FUNCTION_BLOCK T_SafeSr_Tests EXTENDS TcUnit.FB_TestSuite
VAR
    // Test_SetDominantLatch
    group_1 : T_SafeGroup;
    fb_1 : T_SafeSr(group := group_1);
    // Test_UnconnectedResetIsRefused
    group_2 : T_SafeGroup;
    fb_2 : T_SafeSr(group := group_2);
END_VAR

Test_SetDominantLatch();
Test_UnconnectedResetIsRefused();

METHOD PRIVATE Test_SetDominantLatch
TcUnit.TEST(__POUNAME());
// act / assert
group_1(Run := TRUE);
fb_1(Set := TRUE, Reset := TRUE);
AssertEquals_BOOL(Expected := TRUE, Actual := fb_1.SrOut, Message := 'set dominant');
fb_1(Set := FALSE, Reset := TRUE);
AssertEquals_BOOL(Expected := FALSE, Actual := fb_1.SrOut, Message := 'reset');
fb_1(Set := FALSE, Reset := FALSE);
AssertEquals_BOOL(Expected := FALSE, Actual := fb_1.SrOut, Message := 'held');
TEST_FINISHED_NAMED(__POUNAME());
END_METHOD

METHOD PRIVATE Test_UnconnectedResetIsRefused
TcUnit.TEST(__POUNAME());
// arrange / act: Reset is unconnected, which the Safety Editor refuses
group_2(Run := TRUE);
fb_2(Set := TRUE);
group_2(Run := TRUE);
fb_2(Set := TRUE);
// assert
AssertEquals_BOOL(Expected := TRUE, Actual := fb_2.Error, Message := 'configuration error reported');
AssertEquals_BYTE(Expected := TO_BYTE(E_SafeFbState.Error), Actual := fb_2.State, Message := 'state ERROR');
AssertEquals_WORD(Expected := WORD#16#8000, Actual := fb_2.Diag, Message := 'diag bit 15 configuration refused');
AssertEquals_BOOL(Expected := FALSE, Actual := fb_2.SrOut, Message := 'SrOut stays at its safe value');
AssertEquals_BOOL(Expected := TRUE, Actual := group_2.FbErr, Message := 'the group sees an FB error');
// act: ErrAck 0 -> 1 -> 0 does not clear a configuration error
group_2(Run := TRUE, ErrAck := TRUE);
fb_2(Set := TRUE);
group_2(Run := TRUE, ErrAck := TRUE);
fb_2(Set := TRUE);
group_2(Run := TRUE, ErrAck := FALSE);
fb_2(Set := TRUE);
AssertEquals_BOOL(Expected := TRUE, Actual := fb_2.Error, Message := 'error not acknowledged');
AssertEquals_WORD(Expected := WORD#16#8000, Actual := fb_2.Diag, Message := 'diag bit 15 kept');
TEST_FINISHED_NAMED(__POUNAME());
END_METHOD

END_FUNCTION_BLOCK

(* stored: Version 1.1.0.1
   POU T_SafeSr_Tests: Id {1d7ca810-c3c7-5427-960e-46985b1d864e}, SpecialFunc None
   Method Test_SetDominantLatch: Id {0101a96f-fe80-50b6-94a4-1d27727dfa03}
   Method Test_UnconnectedResetIsRefused: Id {4f489207-db0a-4806-8073-86bdcc60f989} *)
